Staubli VAL3: CalToolPos3.pgx

public program CalToolPos3(tool& x_tTool)
  local bool l_bStatus
  local pointRs l_p1
  local pointRs l_p2
  local pointRs l_p3
  local pointRs l_pCenter
  local tool l_t1
  local tool l_t2
  local tool l_t3
begin
  l_bStatus=false
  link(l_pCenter,world)
  //
  l_p1=db:pTeach1
  l_p2=db:pTeach2
  l_p3=db:pTeach3
  call _CalpCircle(l_p1,l_p2,l_p3,l_pCenter,l_bStatus)
  //

  if l_bStatus==true
    l_pCenter.trsf.rx=0
    l_pCenter.trsf.ry=180
    l_pCenter.trsf.rz=0
  else
    call db:hmiAlert("DeviationIsTooLarge","warning")
  endIf
  l_t1.trsf=!l_p1.trsf*l_pCenter.trsf
  l_t2.trsf=!l_p2.trsf*l_pCenter.trsf
  l_t3.trsf=!l_p3.trsf*l_pCenter.trsf
  x_tTool.trsf.x=(l_t1.trsf.x+l_t2.trsf.x+l_t3.trsf.x)/3
  x_tTool.trsf.y=(l_t1.trsf.y+l_t2.trsf.y+l_t3.trsf.y)/3
  x_tTool.trsf.z=0
  x_tTool.trsf.rx=0
  x_tTool.trsf.ry=0
  x_tTool.trsf.rz=0
  call db:hmiAlert("SaveInTool1","info")
end
